{attribute 'enable_dynamic_creation'}
FUNCTION_BLOCK FB_KeyValue IMPLEMENTS I_OtlpValue
VAR_OUTPUT
	pKey: POINTER TO STRING;
	pVal: POINTER TO FB_AnyValue;
END_VAR

(*
	Releases this value and clears the caller's pointer to it: call it as p^.delete(pSelf:=p).
	pSelf is cleared before the value is freed, so the caller never keeps a dangling pointer.
	A pointer to any other object is refused and left untouched, and nothing is released.
*)
METHOD delete : BOOL
VAR_IN_OUT
	pSelf: POINTER TO FB_KeyValue;
END_VAR
VAR
	_pThis: POINTER TO FB_KeyValue;
END_VAR
_pThis := THIS;
IF pSelf <> _pThis THEN
	RETURN;
END_IF

pSelf := 0;
__DELETE(_pThis);
delete := TRUE;
END_METHOD

PROPERTY eType : E_ValueType
GET
eType := E_ValueType.E_KeyValue;
END_GET
END_PROPERTY

//FB_Exit must be implemented explicitly. If there is an implementation, then the
//method is called before the controller removes the code of the function block instance
//(implicit call). The return value is not evaluated.
METHOD FB_Exit: BOOL
VAR_INPUT
    bInCopyCode: BOOL;  // TRUE: the exit method is called in order to leave the instance which will be copied afterwards (online change).  
END_VAR
THIS^.free();
END_METHOD

//FB_Init is always available implicitly and it is used primarily for initialization.
//The return value is not evaluated. For a specific influence, you can also declare the
//methods explicitly and provide additional code there with the standard initialization
//code. You can evaluate the return value.
METHOD FB_Init: BOOL
VAR_INPUT
    bInitRetains: BOOL; // TRUE: the retain variables are initialized (reset warm / reset cold)
    bInCopyCode: BOOL;  // TRUE: the instance will be copied to the copy code afterward (online change)
	pKey: POINTER TO STRING;
	pVal: POINTER TO FB_AnyValue;
END_VAR
(* Validation and allocation are handled by ValueFactory.createKeyValue. The
factory transfers ownership of both pointers only after every step succeeds. *)
THIS^.pKey := pKey;
THIS^.pVal := pVal;
END_METHOD

(* deallocates all data owned by the value without deleting the object itself.*)
METHOD free
IF THIS^.pKey <> 0 THEN
	__DELETE(THIS^.pKey);
	THIS^.pKey := 0;
END_IF
IF THIS^.pVal <> 0 THEN
	THIS^.pVal^.delete(pSelf:=THIS^.pVal);
END_IF
END_METHOD

END_FUNCTION_BLOCK

(* stored: Version 1.1.0.1
   POU FB_KeyValue: Id {8780a23e-cbf3-48bf-8fff-1d17430936ad}, SpecialFunc None
   Method delete: Id {72419ca3-b889-48b2-ba00-e715a127399e}
   Property eType: Id {c2e82dd7-6dca-4765-8d95-f8cdb21c0a06}
   Get Get: Id {2d2213cf-22e8-45af-948d-469cf23853fd}
   Method FB_Exit: Id {3e29dca2-c132-46d7-b434-02454cf38aee}
   Method FB_Init: Id {0ded1b83-877d-444a-a70d-64070bc67700}
   Method free: Id {f43303d8-cb9a-4788-90b7-d0e19760a4b9} *)
